Fanuc KAREL source: KA00149.KL

PROGRAM KA00149
%NOLOCKGROUP
VAR
  SRC: ARRAY[4] OF INTEGER
  DST: ARRAY[4] OF BYTE
BEGIN
  DST = SRC
END KA00149
